Universal Robots PolyScope program: SpeedProg.urp

Program SpeedProg (createdIn=3.0.0 lastSavedIn=3.0.0 directory=/programs installation=default)
Robot Program (runOnlyOnce=true motionType=MoveJ speed=1.047198 acceleration=1.396263 useActiveTCP=false)
  'Program generated by RoboDK v6.0.7 for ABB IRB 120-3/0.6 on XX/XX/XXXX 18:00:00'
  'Using nominal kinematics.'
  'Using Ref. Frame S: p[1.234570, -0.098765, 0.050500, 0.000000, 0.000000, 0.523599]'
  'Using TCP Tool S: p[0.010000, 0.020000, 0.150000, 0.000000, 0.000000, 0.000000]'
  Script: set_tcp(p[0.010000, 0.020000, 0.150000, 0.000000, 0.000000, 0.000000])
  MoveL speed 1 mm/s, acceleration 1200 mm/s^2 (useActiveTCP=true)
    Waypoint Waypoint_1: motionParameters(blendRadius=0); TCP in base x=436.232 y=68.297 z=413.715 mm, rx=0.1383 ry=2.2532 rz=-0.2966 rad; joints [0, -10, 20, 0, 30, 0] deg; flange x=327.703 y=87.801 z=517.836 mm, rx=0.1383 ry=2.2532 rz=-0.2966 rad
  Script: movej([0.000000, -0.174533, 0.349066, 0.000000, 0.523599, 0.000000],1.20000,0.01745,0,0.0000)
  MoveL speed 12 mm/s, acceleration 1200 mm/s^2 (useActiveTCP=true)
    Waypoint Waypoint_2: motionParameters(blendRadius=0.001); TCP in base x=426.318 y=20 z=422.034 mm, rx=0.1383 ry=2.2532 rz=-0.2966 rad; joints [0, -10, 20, 0, 30, 0] deg; flange x=317.789 y=39.504 z=526.155 mm, rx=0.1383 ry=2.2532 rz=-0.2966 rad
  Script: movej([0.349066, -0.174533, 0.349066, 0.000000, 0.523599, 0.000000],1.20000,0.09599,0,0.0000)
  MoveL speed 100 mm/s, acceleration 1200 mm/s^2 (useActiveTCP=true)
    Waypoint Waypoint_3: motionParameters(blendRadius=0.003); TCP in base x=436.232 y=68.297 z=413.715 mm, rx=0.1383 ry=2.2532 rz=-0.2966 rad; joints [0, -10, 20, 0, 30, 0] deg; flange x=327.703 y=87.801 z=517.836 mm, rx=0.1383 ry=2.2532 rz=-0.2966 rad
  Script: movej([0.000000, -0.174533, 0.349066, 0.000000, 0.523599, 0.000000],1.20000,0.34907,0,0.0000)
  MoveL speed 333 mm/s, acceleration 1200 mm/s^2 (useActiveTCP=true)
    Waypoint Waypoint_4: motionParameters(blendRadius=0.004); TCP in base x=426.318 y=20 z=422.034 mm, rx=0.1383 ry=2.2532 rz=-0.2966 rad; joints [0, -10, 20, 0, 30, 0] deg; flange x=317.789 y=39.504 z=526.155 mm, rx=0.1383 ry=2.2532 rz=-0.2966 rad
  Script: movej([0.349066, -0.174533, 0.349066, 0.000000, 0.523599, 0.000000],1.20000,0.78540,0,0.0000)
  MoveL speed 1000 mm/s, acceleration 1200 mm/s^2 (useActiveTCP=true)
    Waypoint Waypoint_5: motionParameters(blendRadius=0.006); TCP in base x=436.232 y=68.297 z=413.715 mm, rx=0.1383 ry=2.2532 rz=-0.2966 rad; joints [0, -10, 20, 0, 30, 0] deg; flange x=327.703 y=87.801 z=517.836 mm, rx=0.1383 ry=2.2532 rz=-0.2966 rad
  Script: movej([0.000000, -0.174533, 0.349066, 0.000000, 0.523599, 0.000000],1.20000,1.57080,0,0.0000)
  MoveL speed 2500 mm/s, acceleration 1200 mm/s^2 (useActiveTCP=true)
    Waypoint Waypoint_6: motionParameters(blendRadius=0.009); TCP in base x=426.318 y=20 z=422.034 mm, rx=0.1383 ry=2.2532 rz=-0.2966 rad; joints [0, -10, 20, 0, 30, 0] deg; flange x=317.789 y=39.504 z=526.155 mm, rx=0.1383 ry=2.2532 rz=-0.2966 rad
  Script: movej([0.349066, -0.174533, 0.349066, 0.000000, 0.523599, 0.000000],1.20000,2.09440,0,0.0000)
  MoveL speed 3000 mm/s, acceleration 1200 mm/s^2 (useActiveTCP=true)
    Waypoint Waypoint_7: motionParameters(blendRadius=0.015); TCP in base x=436.232 y=68.297 z=413.715 mm, rx=0.1383 ry=2.2532 rz=-0.2966 rad; joints [0, -10, 20, 0, 30, 0] deg; flange x=327.703 y=87.801 z=517.836 mm, rx=0.1383 ry=2.2532 rz=-0.2966 rad
  Script: movej([0.000000, -0.174533, 0.349066, 0.000000, 0.523599, 0.000000],1.20000,3.14159,0,0.0000)
  MoveL speed 3000 mm/s, acceleration 1200 mm/s^2 (useActiveTCP=true)
    Waypoint Waypoint_8: motionParameters(blendRadius=0.03); TCP in base x=426.318 y=20 z=422.034 mm, rx=0.1383 ry=2.2532 rz=-0.2966 rad; joints [0, -10, 20, 0, 30, 0] deg; flange x=317.789 y=39.504 z=526.155 mm, rx=0.1383 ry=2.2532 rz=-0.2966 rad
  Script: movej([0.349066, -0.174533, 0.349066, 0.000000, 0.523599, 0.000000],1.20000,3.14159,0,0.0000)
  MoveL speed 1 mm/s, acceleration 1200 mm/s^2 (useActiveTCP=true)
    Waypoint Waypoint_9: motionParameters(blendRadius=0.075); TCP in base x=436.232 y=68.297 z=413.715 mm, rx=0.1383 ry=2.2532 rz=-0.2966 rad; joints [0, -10, 20, 0, 30, 0] deg; flange x=327.703 y=87.801 z=517.836 mm, rx=0.1383 ry=2.2532 rz=-0.2966 rad
  Script: movej([0.000000, -0.174533, 0.349066, 0.000000, 0.523599, 0.000000],1.20000,3.14159,0,0.0000)
  MoveL speed 750 mm/s, acceleration 1200 mm/s^2 (useActiveTCP=true)
    Waypoint Waypoint_10: motionParameters(blendRadius=0.15); TCP in base x=426.318 y=20 z=422.034 mm, rx=0.1383 ry=2.2532 rz=-0.2966 rad; joints [0, -10, 20, 0, 30, 0] deg; flange x=317.789 y=39.504 z=526.155 mm, rx=0.1383 ry=2.2532 rz=-0.2966 rad
  Script: movej([0.349066, -0.174533, 0.349066, 0.000000, 0.523599, 0.000000],1.20000,0.03927,0,0.0000)
  MoveL speed 750 mm/s, acceleration 2000 mm/s^2 (useActiveTCP=true)
    Waypoint Waypoint_11: motionParameters(blendRadius=0.15); TCP in base x=426.318 y=20 z=422.034 mm, rx=0.1383 ry=2.2532 rz=-0.2966 rad; joints [0, -10, 20, 0, 30, 0] deg; flange x=317.789 y=39.504 z=526.155 mm, rx=0.1383 ry=2.2532 rz=-0.2966 rad
